Fanuc KAREL source: kt00184.KL

-- PROVISIONAL review KL for V1013-1; original PC SHA256 775de959b69a4ef41ceb60cb4f90dd709e2c685470df44c5602345e28f309feb
-- Incomplete behavior may be omitted. Consult companion uncertainty JSON. Do not deploy.
PROGRAM KT00184
%NOLOCKGROUP
VAR
  OUT : REAL
-- UNRESOLVED_DECL Y1 type=002018
-- UNRESOLVED_DECL H2 type=002017
BEGIN
  -- UNRESOLVED_PC offsets 5-19; opcodes 2E,22,9D,33,B2
  -- UNRESOLVED_PC offsets 24-38; opcodes 2E,22,9D,33,B4
  -- UNRESOLVED_PC offsets 43-69; opcodes 22,9D,33,B1,22,9D,33,B3,56,64,23
  -- UNRESOLVED_PC offsets 74-78; opcodes 7F
END KT00184
